(* IEC 61131-3 sources: plc-vscode/tests/st/test-ready/trust-platform/examples/OSCAT/chiller_temperature_pid/non-oop/src, 3 files *)

(* ---- Configuration.st ---- *)
CONFIGURATION ChillerTemperaturePidClassicConfiguration
RESOURCE Cpu0 ON PLC
    TASK MainTask (INTERVAL := T#100ms, PRIORITY := 1);
    PROGRAM Main WITH MainTask : Main;
END_RESOURCE
END_CONFIGURATION

(* ---- Main.st ---- *)
PROGRAM Main
VAR
    TemperatureConversion : TEMPERATURE;
    ChillerController : CTRL_PID;
    ReturnTemperatureCelsius : REAL := REAL#12.0;
    ReturnTemperatureKelvin : REAL;
    ValveCommandPercent : REAL;
END_VAR

TemperatureConversion(C := ReturnTemperatureCelsius);
ReturnTemperatureKelvin := TemperatureConversion.YK;
ChillerController(
    ACT := ReturnTemperatureCelsius,
    SET_POINT := REAL#7.0,
    SUP := REAL#0.0,
    OFS := REAL#0.0,
    M_I := REAL#45.0,
    MAN := TRUE,
    RST := FALSE,
    KP := REAL#2.0,
    TN := REAL#1.0,
    TV := REAL#0.0,
    LL := REAL#0.0,
    LH := REAL#100.0
);
ValveCommandPercent := ChillerController.Y;
END_PROGRAM

(* ---- Tests.st ---- *)
TEST_PROGRAM ChillerTemperaturePidClassicConvertsAndControls
VAR
    TemperatureConversion : TEMPERATURE;
    ChillerController : CTRL_PID;
END_VAR

TemperatureConversion(C := REAL#12.0);
ChillerController(
    ACT := REAL#12.0,
    SET_POINT := REAL#7.0,
    SUP := REAL#0.0,
    OFS := REAL#0.0,
    M_I := REAL#45.0,
    MAN := TRUE,
    RST := FALSE,
    KP := REAL#2.0,
    TN := REAL#1.0,
    TV := REAL#0.0,
    LL := REAL#0.0,
    LH := REAL#100.0
);

ASSERT_NEAR(EXPECTED := REAL#285.15, ACTUAL := TemperatureConversion.YK, DELTA := REAL#0.01);
ASSERT_NEAR(EXPECTED := REAL#45.0, ACTUAL := ChillerController.Y, DELTA := REAL#0.001);
END_TEST_PROGRAM
